Fanuc KAREL source: KA00190.KL

PROGRAM KA00190
%NOLOCKGROUP
VAR
  SRC: ARRAY[4] OF SHORT
  DST: ARRAY[4] OF INTEGER
BEGIN
  DST = SRC
END KA00190
